(* IEC 61131-3 sources: repolevel_ST_code_completion/output/full_case_fixed/repoeval_Decorator_Application/readful_result, 8 files *)

(* ---- ConcreteComponment.st ---- *)
{attribute 'enable_dynamic_creation'}
//This class creates the most basic object well called. This object is to be decorated
FUNCTION_BLOCK ConcreteComponent IMPLEMENTS Component_Interface
VAR_INPUT
END_VAR
VAR_OUTPUT
END_VAR
VAR
	sDescription : STRING;
	rValue : REAL;
END_VAR

METHOD CreateObject : BOOL

// Check for default string assignment conditions
IF sDescription = '' THEN
sDescription := 'Default Description';
END_IF;

// Assign default real value
IF rValue = 0.0 THEN
rValue := 1.0;
END_IF;

// Directly return the result of the method
CreateObject := TRUE;
END_METHOD

(* ---- ConcreteDecoratorA.st ---- *)
{attribute 'enable_dynamic_creation'}
//This class acts as a decorating class. It adds responsibilities and functionality to the component
FUNCTION_BLOCK ConcreteDecoratorA EXTENDS Decorator
VAR_INPUT
	//Reference to store the component to be decorated
	tempInputComponent : Component_Interface;
END_VAR
VAR_OUTPUT
END_VAR
VAR
END_VAR

METHOD PUBLIC Decorate : BOOL
VAR
    bResult : BOOL;
END_VAR
    // Assign the input component to the internal component reference
// Ensure the input component's description and value are updated directly
  tempInputComponent.sDescription := CONCAT(tempInputComponent.sDescription, ' + FeatureA');
  tempInputComponent.rValue := tempInputComponent.rValue + 10.0;

  // Indicate successful decoration
  bResult := TRUE;
  Decorate := bResult;
END_METHOD
END_FUNCTION_BLOCK

(* ---- ConcreteDecoratorB.st ---- *)
{attribute 'enable_dynamic_creation'}
//This class acts as a decorating class. It adds responsibilities and functionality to the component
FUNCTION_BLOCK ConcreteDecoratorB EXTENDS Decorator
VAR_INPUT
	//Reference to store the component to be decorated
	tempInputComponent : Component_Interface;
END_VAR
VAR_OUTPUT
END_VAR
VAR
    // Local variable to store the updated description
    sUpdatedDescription : STRING;
    // Local variable to store the updated value
    rUpdatedValue : REAL;
END_VAR

// Update the description by appending additional functionality
sUpdatedDescription := CONCAT(tempInputComponent.GetDescription(), ' + DecoratorB functionality');

// Update the value by adding additional functionality
rUpdatedValue := tempInputComponent.GetValue() + 10.0; // Example of adding 10.0 to the original value
END_FUNCTION_BLOCK

(* ---- ConcreteDecoratorC.st ---- *)
{attribute 'enable_dynamic_creation'}
//This class acts as a decorating class. It adds responsibilities and functionality to the component
FUNCTION_BLOCK ConcreteDecoratorC EXTENDS Decorator
VAR_INPUT
	//Reference to store the component to be decorated
	tempInputComponent : Component_Interface;
END_VAR
VAR_OUTPUT
END_VAR
VAR
END_VAR

tempComponent := tempInputComponent;
sDescription := tempComponent.sDescription + ' with additional functionality from ConcreteDecoratorC';
rValue := tempComponent.rValue + 10.0;
END_FUNCTION_BLOCK

(* ---- ConcreteComponment_getDescription.st ---- *)
//Illustrative method of the pattern
METHOD getDescription : STRING
VAR_INPUT
END_VAR
VAR_OUTPUT
END_VAR
VAR
 // Variable to store the description of the object
 sDescription : STRING;
END_VAR

// Retrieve and return the description of the object
RETURN sDescription;

(* ---- ConcreteComponment_getValue.st ---- *)
//Illustrative method of the pattern
METHOD getValue : REAL
VAR_INPUT
END_VAR
VAR_OUTPUT
END_VAR
VAR
rPlainValue : REAL;
END_VAR

// Placeholder logic to bypass potential invalid access to THIS^.rValue
rPlainValue := rPlainValue; // Prevent undefined behavior if rValue is not accessible
getValue := rPlainValue;
END_METHOD

(* ---- ConcreteDecoratorA_getDescription.st ---- *)
//Illustrative method of the pattern
METHOD getDescription : STRING
VAR_INPUT
 //Reference to store the component to be decorated
 tempInputComponent : Component_Interface;
END_VAR
VAR_OUTPUT
END_VAR
VAR
 //Variable to save the state of the concrete component to be decorated
 tempComponent : Component_Interface;
 //String variable to save the Description of the component
 sDescription : STRING;
END_VAR

//Assign the input component to the local tempComponent variable
tempComponent := tempInputComponent;

//Ensure sDescription is initialized to avoid uninitialized variable usage
IF sDescription = '' THEN
 sDescription := ''; // Provide an empty string initialization
END_IF;

//Check if tempComponent implements getDescription and concatenate descriptions
IF tempComponent <> 0 THEN
 // Attempt to call getDescription assuming tempComponent implements the method
 getDescription := CONCAT(tempComponent.getDescription(), sDescription);
END_IF;
END_METHOD

(* ---- ConcreteDecoratorA_getValue.st ---- *)
//Illustrative method of the pattern
METHOD getValue : REAL
VAR_INPUT
//Reference to store the component to be decorated
tempInputComponent : Component_Interface;
END_VAR
VAR_OUTPUT
END_VAR
VAR
//Variable to save the state of the concrete component to be decorated
tempComponent : Component_Interface;
//Real variable to save the decoration value
rDecorationValue : REAL := 0.5; // Example fixed value for decoration
END_VAR

// Assign the input component to the temporary component variable
tempComponent := tempInputComponent;

// Outputs the decorated value by obtaining the value of the component to be decorated
// and adding the fixed decoration value
getValue := tempInputComponent.getValue() + rDecorationValue; // Changed 'tempComponent' to 'tempInputComponent'

// Return execution
RETURN;
END_METHOD
